(* IEC 61131-3 sources: teller/JD_Teller_LC2_V11/Network/LseRtkMain, 1 file *)

(* ---- ONE_LseRtkMain_Table.st ---- *)
#define OBJECTS_CONFIG

FUNCTION GLOBAL TAB ONE_LseRtkMain
-1$UINT, 0$UINT,
0$UINT, 0$UINT,

24$UDINT,
TO_UDINT(3788417926), "_Global", 0$UINT, 12$UINT, 0$UINT,
TO_UDINT(2996404079), "_LimitMax", 0$UINT, 1$UINT, 1$UINT,
TO_UDINT(2392080438), "_LimitMin", 0$UINT, 1$UINT, 1$UINT,
TO_UDINT(1552551876), "_Lse", 0$UINT, 95$UINT, 1$UINT,
TO_UDINT(2980745877), "_MyIO", 0$UINT, 3$UINT, 0$UINT,
TO_UDINT(3599188277), "_Screen", 0$UINT, 2$UINT, 1$UINT,
TO_UDINT(3931827689), "_SysDateTime", 0$UINT, 5$UINT, 1$UINT,
TO_UDINT(3192771746), "_XAccess", 0$UINT, 1$UINT, 1$UINT,
TO_UDINT(3255080645), "ActScreenWindow", 0$UINT, 0$UINT, 1$UINT,
TO_UDINT(2897291062), "ASCII_BIN", 1$UINT, 20$UINT, 1$UINT,
TO_UDINT(3502790066), "Count_To", 0$UINT, 0$UINT, 1$UINT,
TO_UDINT(809080914), "LoadSaveData", 1$UINT, 0$UINT, 1$UINT,
TO_UDINT(2276934072), "Merker", 1$UINT, 0$UINT, 2$UINT,
TO_UDINT(2225119864), "MerkerEx", 1$UINT, 18$UINT, 22$UINT,
TO_UDINT(311276651), "OperatorLogIn_Teller", 1$UINT, 0$UINT, 1$UINT,
TO_UDINT(1903583397), "Ram", 1$UINT, 3$UINT, 5$UINT,
TO_UDINT(1260770215), "SetPassword", 0$UINT, 0$UINT, 3$UINT,
TO_UDINT(1850111279), "String", 1$UINT, 10$UINT, 22$UINT,
TO_UDINT(2898603620), "StringInternal", 1$UINT, 70$UINT, 0$UINT,
TO_UDINT(2580220589), "Summertime_Selector", 0$UINT, 0$UINT, 1$UINT,
TO_UDINT(4036227488), "SV_Help", 0$UINT, 0$UINT, 1$UINT,
TO_UDINT(74052286), "TerminalControl", 0$UINT, 0$UINT, 1$UINT,
TO_UDINT(2675810274), "Timeconvert", 0$UINT, 0$UINT, 1$UINT,
TO_UDINT(3232495061), "VirtualBaseInit", 1$UINT, 3$UINT, 0$UINT,

_NO_ATTR, TO_UDINT(2623093263), "LIMITMAX",

_NO_ATTR, TO_UDINT(2689860950), "LIMITMIN",

_NO_ATTR, TO_UDINT(299963966), "LSE",

_NO_ATTR, TO_UDINT(2730400835), "_SCREEN0",

_NO_ATTR, TO_UDINT(3035062039), "SYSDATETIME",

_NO_ATTR, TO_UDINT(3799848273), "XACCESS0",

_NO_ATTR, TO_UDINT(1745935646), "ACTSCREENWINDOW1",

1$UINT, TO_UDINT(2522576343), "OPERATORLOGIN1\ASCII_BIN1",

_NO_ATTR, TO_UDINT(2791568706), "COUNT_TO1",

_NO_ATTR, TO_UDINT(109700855), "LOADSAVEDATA1",

_NO_ATTR, TO_UDINT(1180982051), "INSERTLOCK",
_NO_ATTR, TO_UDINT(49391923), "SHIFTLOCK",

1$UINT, TO_UDINT(365676125), "OPERATORLOGIN1\OP01_NAME\MERKEREX0",
1$UINT, TO_UDINT(3330497326), "OPERATORLOGIN1\OP01_WW\MERKEREX0",
1$UINT, TO_UDINT(1006858927), "OPERATORLOGIN1\OP02_NAME\MERKEREX0",
1$UINT, TO_UDINT(3135405813), "OPERATORLOGIN1\OP02_WW\MERKEREX0",
1$UINT, TO_UDINT(2456544062), "OPERATORLOGIN1\OP03_NAME\MERKEREX0",
1$UINT, TO_UDINT(669884291), "OPERATORLOGIN1\OP03_WW\MERKEREX0",
1$UINT, TO_UDINT(1871846219), "OPERATORLOGIN1\OP04_NAME\MERKEREX0",
1$UINT, TO_UDINT(1109407043), "OPERATORLOGIN1\OP04_WW\MERKEREX0",
1$UINT, TO_UDINT(3254422234), "OPERATORLOGIN1\OP05_NAME\MERKEREX0",
1$UINT, TO_UDINT(3744453685), "OPERATORLOGIN1\OP05_WW\MERKEREX0",
1$UINT, TO_UDINT(3895606824), "OPERATORLOGIN1\OP06_NAME\MERKEREX0",
1$UINT, TO_UDINT(2739859950), "OPERATORLOGIN1\OP06_WW\MERKEREX0",
1$UINT, TO_UDINT(1180348345), "OPERATORLOGIN1\OP07_NAME\MERKEREX0",
1$UINT, TO_UDINT(1044451480), "OPERATORLOGIN1\OP07_WW\MERKEREX0",
1$UINT, TO_UDINT(3367028867), "OPERATORLOGIN1\OP08_NAME\MERKEREX0",
1$UINT, TO_UDINT(1758831726), "OPERATORLOGIN1\OP08_WW\MERKEREX0",
1$UINT, TO_UDINT(1725454610), "OPERATORLOGIN1\OP09_NAME\MERKEREX0",
1$UINT, TO_UDINT(4124722456), "OPERATORLOGIN1\OP09_WW\MERKEREX0",
1$UINT, TO_UDINT(1007000719), "OPERATORLOGIN1\OP10_NAME\MERKEREX0",
1$UINT, TO_UDINT(3799474608), "OPERATORLOGIN1\OP10_WW\MERKEREX0",
1$UINT, TO_UDINT(856832036), "OPERATORLOGIN1\OPERATOR_SELECTED\MERKEREX0",
1$UINT, TO_UDINT(608268224), "OPERATORLOGIN1\WW_INVOER\MERKEREX0",

_NO_ATTR, TO_UDINT(3114945658), "OPERATORLOGIN1",

1$UINT, TO_UDINT(1119588755), "SYSDATETIME\SUMMERTIME",
1$UINT, TO_UDINT(440852310), "XACCESS0\RAM0",
1$UINT, TO_UDINT(1833037760), "XACCESS0\RAM1",
1$UINT, TO_UDINT(4098408058), "XACCESS0\RAM2",
1$UINT, TO_UDINT(2203029228), "XACCESS0\RAM3",

_NO_ATTR, TO_UDINT(3408264239), "SETPASSWORD1",
_NO_ATTR, TO_UDINT(1378659733), "SETPASSWORD2",
_NO_ATTR, TO_UDINT(623615235), "SETPASSWORD3",

1$UINT, TO_UDINT(3623239739), "OPERATORLOGIN1\OP01_NAME",
1$UINT, TO_UDINT(1286520628), "OPERATORLOGIN1\OP01_WW",
1$UINT, TO_UDINT(1365389973), "OPERATORLOGIN1\OP02_NAME",
1$UINT, TO_UDINT(1578832090), "OPERATORLOGIN1\OP02_WW",
1$UINT, TO_UDINT(2587812144), "OPERATORLOGIN1\OP03_NAME",
1$UINT, TO_UDINT(3869734847), "OPERATORLOGIN1\OP03_WW",
1$UINT, TO_UDINT(2268844424), "OPERATORLOGIN1\OP04_NAME",
1$UINT, TO_UDINT(2070957830), "OPERATORLOGIN1\OP04_WW",
1$UINT, TO_UDINT(1281819181), "OPERATORLOGIN1\OP05_NAME",
1$UINT, TO_UDINT(3284936803), "OPERATORLOGIN1\OP05_WW",
1$UINT, TO_UDINT(3404951683), "OPERATORLOGIN1\OP06_NAME",
1$UINT, TO_UDINT(3514402701), "OPERATORLOGIN1\OP06_WW",
1$UINT, TO_UDINT(28287782), "OPERATORLOGIN1\OP07_NAME",
1$UINT, TO_UDINT(1774575848), "OPERATORLOGIN1\OP07_WW",
1$UINT, TO_UDINT(4042854899), "OPERATORLOGIN1\OP08_NAME",
1$UINT, TO_UDINT(833024190), "OPERATORLOGIN1\OP08_WW",
1$UINT, TO_UDINT(1000718934), "OPERATORLOGIN1\OP09_NAME",
1$UINT, TO_UDINT(2300221403), "OPERATORLOGIN1\OP09_WW",
1$UINT, TO_UDINT(3135084586), "OPERATORLOGIN1\OP10_NAME",
1$UINT, TO_UDINT(3379753441), "OPERATORLOGIN1\OP10_WW",
1$UINT, TO_UDINT(3938195579), "OPERATORLOGIN1\OPERATOR_SELECTED",
1$UINT, TO_UDINT(3642620268), "OPERATORLOGIN1\WW_INVOER",

_NO_ATTR, TO_UDINT(723713000), "SUMMERTIME_SELECTOR1",

_NO_ATTR, TO_UDINT(1442504622), "SV_HELP1",

_NO_ATTR, TO_UDINT(2936084686), "TERMINALCONTROL1",

_NO_ATTR, TO_UDINT(3443986812), "TIMECONVERT1",

//Internal connections
0$UDINT,
50$UDINT,
TO_UDINT(4), "SummerTime", TO_UDINT(35),
TO_UDINT(5), "Ram0", TO_UDINT(36),
TO_UDINT(5), "Ram1", TO_UDINT(37),
TO_UDINT(5), "Ram2", TO_UDINT(38),
TO_UDINT(5), "Ram3", TO_UDINT(39),
TO_UDINT(34), "Op10_Name", TO_UDINT(61),
TO_UDINT(34), "Op10_WW", TO_UDINT(62),
TO_UDINT(34), "Op01_Name", TO_UDINT(43),
TO_UDINT(34), "Op01_WW", TO_UDINT(44),
TO_UDINT(34), "Op02_Name", TO_UDINT(45),
TO_UDINT(34), "Op02_WW", TO_UDINT(46),
TO_UDINT(34), "Op03_Name", TO_UDINT(47),
TO_UDINT(34), "Op03_WW", TO_UDINT(48),
TO_UDINT(34), "Op04_Name", TO_UDINT(49),
TO_UDINT(34), "Op04_WW", TO_UDINT(50),
TO_UDINT(34), "Op05_Name", TO_UDINT(51),
TO_UDINT(34), "Op05_WW", TO_UDINT(52),
TO_UDINT(34), "Op06_Name", TO_UDINT(53),
TO_UDINT(34), "Op06_WW", TO_UDINT(54),
TO_UDINT(34), "Op07_Name", TO_UDINT(55),
TO_UDINT(34), "Op07_WW", TO_UDINT(56),
TO_UDINT(34), "Op08_Name", TO_UDINT(57),
TO_UDINT(34), "Op08_WW", TO_UDINT(58),
TO_UDINT(34), "Op09_Name", TO_UDINT(59),
TO_UDINT(34), "Op09_WW", TO_UDINT(60),
TO_UDINT(34), "WW_Invoer", TO_UDINT(64),
TO_UDINT(34), "Operator_Selected", TO_UDINT(63),
TO_UDINT(34), "ASCII_BIN1", TO_UDINT(7),
TO_UDINT(43), "MerkerEx0", TO_UDINT(12),
TO_UDINT(44), "MerkerEx0", TO_UDINT(13),
TO_UDINT(45), "MerkerEx0", TO_UDINT(14),
TO_UDINT(46), "MerkerEx0", TO_UDINT(15),
TO_UDINT(47), "MerkerEx0", TO_UDINT(16),
TO_UDINT(48), "MerkerEx0", TO_UDINT(17),
TO_UDINT(49), "MerkerEx0", TO_UDINT(18),
TO_UDINT(50), "MerkerEx0", TO_UDINT(19),
TO_UDINT(51), "MerkerEx0", TO_UDINT(20),
TO_UDINT(52), "MerkerEx0", TO_UDINT(21),
TO_UDINT(53), "MerkerEx0", TO_UDINT(22),
TO_UDINT(54), "MerkerEx0", TO_UDINT(23),
TO_UDINT(55), "MerkerEx0", TO_UDINT(24),
TO_UDINT(56), "MerkerEx0", TO_UDINT(25),
TO_UDINT(57), "MerkerEx0", TO_UDINT(26),
TO_UDINT(58), "MerkerEx0", TO_UDINT(27),
TO_UDINT(59), "MerkerEx0", TO_UDINT(28),
TO_UDINT(60), "MerkerEx0", TO_UDINT(29),
TO_UDINT(61), "MerkerEx0", TO_UDINT(30),
TO_UDINT(62), "MerkerEx0", TO_UDINT(31),
TO_UDINT(63), "MerkerEx0", TO_UDINT(32),
TO_UDINT(64), "MerkerEx0", TO_UDINT(33),
0$UDINT,
36$UDINT,
TO_UDINT(0), "Lse", TO_UDINT(2), "Lse",
TO_UDINT(1), "Lse", TO_UDINT(2), "Lse",
TO_UDINT(3), "Lse", TO_UDINT(2), "Lse",
TO_UDINT(4), "DoSummerTime", TO_UDINT(65), "SetRegion",
TO_UDINT(5), "Lse", TO_UDINT(2), "Lse",
TO_UDINT(6), "Lse", TO_UDINT(2), "Lse",
TO_UDINT(34), "inlogNiveau", TO_UDINT(5), "Level",
TO_UDINT(34), "c_SysDateTime", TO_UDINT(4), "SysDate",
TO_UDINT(34), "objLoadSaveData", TO_UDINT(9), "ClassSvr",
TO_UDINT(40), "ActKey", TO_UDINT(5), "Key1",
TO_UDINT(41), "ActKey", TO_UDINT(5), "Key2",
TO_UDINT(42), "ActKey", TO_UDINT(5), "Key3",
TO_UDINT(43), "DataBuffer", TO_UDINT(12), "m_udLength",
TO_UDINT(44), "DataBuffer", TO_UDINT(13), "m_udLength",
TO_UDINT(45), "DataBuffer", TO_UDINT(14), "m_udLength",
TO_UDINT(46), "DataBuffer", TO_UDINT(15), "m_udLength",
TO_UDINT(47), "DataBuffer", TO_UDINT(16), "m_udLength",
TO_UDINT(48), "DataBuffer", TO_UDINT(17), "m_udLength",
TO_UDINT(49), "DataBuffer", TO_UDINT(18), "m_udLength",
TO_UDINT(50), "DataBuffer", TO_UDINT(19), "m_udLength",
TO_UDINT(51), "DataBuffer", TO_UDINT(20), "m_udLength",
TO_UDINT(52), "DataBuffer", TO_UDINT(21), "m_udLength",
TO_UDINT(53), "DataBuffer", TO_UDINT(22), "m_udLength",
TO_UDINT(54), "DataBuffer", TO_UDINT(23), "m_udLength",
TO_UDINT(55), "DataBuffer", TO_UDINT(24), "m_udLength",
TO_UDINT(56), "DataBuffer", TO_UDINT(25), "m_udLength",
TO_UDINT(57), "DataBuffer", TO_UDINT(26), "m_udLength",
TO_UDINT(58), "DataBuffer", TO_UDINT(27), "m_udLength",
TO_UDINT(59), "DataBuffer", TO_UDINT(28), "m_udLength",
TO_UDINT(60), "DataBuffer", TO_UDINT(29), "m_udLength",
TO_UDINT(61), "DataBuffer", TO_UDINT(30), "m_udLength",
TO_UDINT(62), "DataBuffer", TO_UDINT(31), "m_udLength",
TO_UDINT(63), "DataBuffer", TO_UDINT(32), "m_udLength",
TO_UDINT(64), "DataBuffer", TO_UDINT(33), "m_udLength",
TO_UDINT(67), "Lse", TO_UDINT(2), "Lse",
TO_UDINT(68), "Milisecs", TO_UDINT(5), "TimeOut",

//Initialization values
0$UDINT,
55$UDINT,
TO_UDINT(2), "SeekAlgorithm", TO_UDINT(1),//|LseRtkMain.Lse.SeekAlgorithm;
TO_UDINT(3), "No", TO_UDINT(0),//|LseRtkMain._Screen0.No;
TO_UDINT(3), "ImA", TO_UDINT(IMA_PICTURE),//|LseRtkMain._Screen0.ImA;
TO_UDINT(4), "DoSummerTime", TO_UDINT(0),//|LseRtkMain.SysDateTime.DoSummerTime;
TO_UDINT(12), "ThreadSafe", TO_UDINT(0),//|LseRtkMain.Op01_Name\OperatorLogIn1\MerkerEx0.ThreadSafe;
TO_UDINT(13), "ThreadSafe", TO_UDINT(0),//|LseRtkMain.Op01_WW\OperatorLogIn1\MerkerEx0.ThreadSafe;
TO_UDINT(14), "ThreadSafe", TO_UDINT(0),//|LseRtkMain.Op02_Name\OperatorLogIn1\MerkerEx0.ThreadSafe;
TO_UDINT(15), "ThreadSafe", TO_UDINT(0),//|LseRtkMain.Op02_WW\OperatorLogIn1\MerkerEx0.ThreadSafe;
TO_UDINT(16), "ThreadSafe", TO_UDINT(0),//|LseRtkMain.Op03_Name\OperatorLogIn1\MerkerEx0.ThreadSafe;
TO_UDINT(17), "ThreadSafe", TO_UDINT(0),//|LseRtkMain.Op03_WW\OperatorLogIn1\MerkerEx0.ThreadSafe;
TO_UDINT(18), "ThreadSafe", TO_UDINT(0),//|LseRtkMain.Op04_Name\OperatorLogIn1\MerkerEx0.ThreadSafe;
TO_UDINT(19), "ThreadSafe", TO_UDINT(0),//|LseRtkMain.Op04_WW\OperatorLogIn1\MerkerEx0.ThreadSafe;
TO_UDINT(20), "ThreadSafe", TO_UDINT(0),//|LseRtkMain.Op05_Name\OperatorLogIn1\MerkerEx0.ThreadSafe;
TO_UDINT(21), "ThreadSafe", TO_UDINT(0),//|LseRtkMain.Op05_WW\OperatorLogIn1\MerkerEx0.ThreadSafe;
TO_UDINT(22), "ThreadSafe", TO_UDINT(0),//|LseRtkMain.Op06_Name\OperatorLogIn1\MerkerEx0.ThreadSafe;
TO_UDINT(23), "ThreadSafe", TO_UDINT(0),//|LseRtkMain.Op06_WW\OperatorLogIn1\MerkerEx0.ThreadSafe;
TO_UDINT(24), "ThreadSafe", TO_UDINT(0),//|LseRtkMain.Op07_Name\OperatorLogIn1\MerkerEx0.ThreadSafe;
TO_UDINT(25), "ThreadSafe", TO_UDINT(0),//|LseRtkMain.Op07_WW\OperatorLogIn1\MerkerEx0.ThreadSafe;
TO_UDINT(26), "ThreadSafe", TO_UDINT(0),//|LseRtkMain.Op08_Name\OperatorLogIn1\MerkerEx0.ThreadSafe;
TO_UDINT(27), "ThreadSafe", TO_UDINT(0),//|LseRtkMain.Op08_WW\OperatorLogIn1\MerkerEx0.ThreadSafe;
TO_UDINT(28), "ThreadSafe", TO_UDINT(0),//|LseRtkMain.Op09_Name\OperatorLogIn1\MerkerEx0.ThreadSafe;
TO_UDINT(29), "ThreadSafe", TO_UDINT(0),//|LseRtkMain.Op09_WW\OperatorLogIn1\MerkerEx0.ThreadSafe;
TO_UDINT(30), "ThreadSafe", TO_UDINT(0),//|LseRtkMain.Op10_Name\OperatorLogIn1\MerkerEx0.ThreadSafe;
TO_UDINT(31), "ThreadSafe", TO_UDINT(0),//|LseRtkMain.Op10_WW\OperatorLogIn1\MerkerEx0.ThreadSafe;
TO_UDINT(32), "ThreadSafe", TO_UDINT(0),//|LseRtkMain.Operator_Selected\OperatorLogIn1\MerkerEx0.ThreadSafe;
TO_UDINT(33), "ThreadSafe", TO_UDINT(0),//|LseRtkMain.WW_Invoer\OperatorLogIn1\MerkerEx0.ThreadSafe;
TO_UDINT(40), "Always", TO_UDINT(1),//|LseRtkMain.SetPassword1.Always;
TO_UDINT(40), "PreSetKey", TO_UDINT(123),//|LseRtkMain.SetPassword1.PreSetKey;
TO_UDINT(41), "Always", TO_UDINT(1),//|LseRtkMain.SetPassword2.Always;
TO_UDINT(41), "PreSetKey", TO_UDINT(416477),//|LseRtkMain.SetPassword2.PreSetKey;
TO_UDINT(42), "Always", TO_UDINT(1),//|LseRtkMain.SetPassword3.Always;
TO_UDINT(42), "PreSetKey", TO_UDINT(552125),//|LseRtkMain.SetPassword3.PreSetKey;
TO_UDINT(43), "SingleRealloc", TO_UDINT(1),//|LseRtkMain.OperatorLogIn1\Op01_Name.SingleRealloc;
TO_UDINT(44), "SingleRealloc", TO_UDINT(1),//|LseRtkMain.OperatorLogIn1\Op01_WW.SingleRealloc;
TO_UDINT(45), "SingleRealloc", TO_UDINT(1),//|LseRtkMain.OperatorLogIn1\Op02_Name.SingleRealloc;
TO_UDINT(46), "SingleRealloc", TO_UDINT(1),//|LseRtkMain.OperatorLogIn1\Op02_WW.SingleRealloc;
TO_UDINT(47), "SingleRealloc", TO_UDINT(1),//|LseRtkMain.OperatorLogIn1\Op03_Name.SingleRealloc;
TO_UDINT(48), "SingleRealloc", TO_UDINT(1),//|LseRtkMain.OperatorLogIn1\Op03_WW.SingleRealloc;
TO_UDINT(49), "SingleRealloc", TO_UDINT(1),//|LseRtkMain.OperatorLogIn1\Op04_Name.SingleRealloc;
TO_UDINT(50), "SingleRealloc", TO_UDINT(1),//|LseRtkMain.OperatorLogIn1\Op04_WW.SingleRealloc;
TO_UDINT(51), "SingleRealloc", TO_UDINT(1),//|LseRtkMain.OperatorLogIn1\Op05_Name.SingleRealloc;
TO_UDINT(52), "SingleRealloc", TO_UDINT(1),//|LseRtkMain.OperatorLogIn1\Op05_WW.SingleRealloc;
TO_UDINT(53), "SingleRealloc", TO_UDINT(1),//|LseRtkMain.OperatorLogIn1\Op06_Name.SingleRealloc;
TO_UDINT(54), "SingleRealloc", TO_UDINT(1),//|LseRtkMain.OperatorLogIn1\Op06_WW.SingleRealloc;
TO_UDINT(55), "SingleRealloc", TO_UDINT(1),//|LseRtkMain.OperatorLogIn1\Op07_Name.SingleRealloc;
TO_UDINT(56), "SingleRealloc", TO_UDINT(1),//|LseRtkMain.OperatorLogIn1\Op07_WW.SingleRealloc;
TO_UDINT(57), "SingleRealloc", TO_UDINT(1),//|LseRtkMain.OperatorLogIn1\Op08_Name.SingleRealloc;
TO_UDINT(58), "SingleRealloc", TO_UDINT(1),//|LseRtkMain.OperatorLogIn1\Op08_WW.SingleRealloc;
TO_UDINT(59), "SingleRealloc", TO_UDINT(1),//|LseRtkMain.OperatorLogIn1\Op09_Name.SingleRealloc;
TO_UDINT(60), "SingleRealloc", TO_UDINT(1),//|LseRtkMain.OperatorLogIn1\Op09_WW.SingleRealloc;
TO_UDINT(61), "SingleRealloc", TO_UDINT(1),//|LseRtkMain.OperatorLogIn1\Op10_Name.SingleRealloc;
TO_UDINT(62), "SingleRealloc", TO_UDINT(1),//|LseRtkMain.OperatorLogIn1\Op10_WW.SingleRealloc;
TO_UDINT(63), "SingleRealloc", TO_UDINT(1),//|LseRtkMain.OperatorLogIn1\Operator_Selected.SingleRealloc;
TO_UDINT(64), "SingleRealloc", TO_UDINT(1),//|LseRtkMain.OperatorLogIn1\WW_Invoer.SingleRealloc;
TO_UDINT(67), "cNextScreen", TO_UDINT(0),//|LseRtkMain.TerminalControl1.cNextScreen;

//Symbolic initialization values
0$UDINT,
0$UDINT,

//Initialization of string values
0$UDINT,
0$UDINT,

//Configuration of tasks (RealTime, Cyclic, Background)
0$UDINT,
0$UDINT,

0$UDINT,
1$UDINT,
TO_UDINT(67), (cCT)$UDINT, 4194305$DINT, 	//TERMINALCONTROL1

0$UDINT,
6$UDINT,
TO_UDINT(2), (-1)$UDINT, 4194305$DINT, 	//LSE
TO_UDINT(4), (250)$UDINT, 4194305$DINT, 	//SYSDATETIME
TO_UDINT(8), (250)$UDINT, 4194305$DINT, 	//COUNT_TO1
TO_UDINT(34), (100)$UDINT, 4194305$DINT, 	//OPERATORLOGIN1
TO_UDINT(65), (250)$UDINT, 4194305$DINT, 	//SUMMERTIME_SELECTOR1
TO_UDINT(68), (100)$UDINT, 4194305$DINT, 	//TIMECONVERT1

//External connections
0$UDINT,
3$UDINT,
TO_UDINT(34), "c_NewFileString", C_DIR, TO_UDINT(738229999), "ToolLight1\NewFileString","Data",
TO_UDINT(34), "c_SelectedFileString", C_DIR, TO_UDINT(639965759), "ToolLight1\FileHandling\toOpenFileStr","Data",
TO_UDINT(34), "c_StringPath", C_DIR, TO_UDINT(107307615), "ToolLight1\FileHandling\PathString","Data",

//Magic internal connections
0$UDINT,
0$UDINT,

//Configuration of timeslots of tasks (RealTime, Cyclic)
#ifdef __LSLLDR_TIMESLOTS__
0$UDINT,
0$UDINT,

0$UDINT,
0$UDINT,

#endif //__LSLLDR_TIMESLOTS__

//MultiMaster connections
#ifdef __LSLLDR_MULTIMASTER__
0$UDINT,
0$UDINT,
#endif //__LSLLDR_MULTIMASTER__

END_FUNCTION
